ABB RobotStudio station: robot-studio-project.rspag

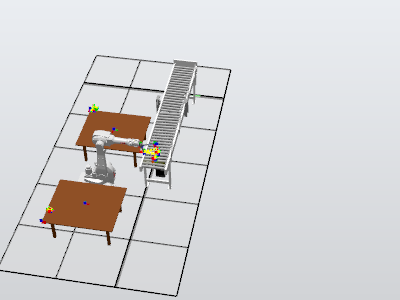
--- station ---
Station FinalConveyor (saved by RobotStudio 24.1.10693.0)
Controller IRB1600_6_145, task T_ROB1: task frame (RAPID world) sits at (2850, -850, 0) mm, rotated rx 0 ry 0 rz 90 deg in the station
Controller IRB1600_6_145
  mechanical unit ROB_1: IRB1600_6_145__03, 6 joints, base frame (0, 0, 0) mm
Layout (positions relative to the parent item):
  - big cube [part], size 200 x 200 x 200 mm
  - small cube [part], size 100 x 100 x 100 mm
  - Conveyor [smart component]
      signals: DI start_or_resume, DO cube_ready, DO cube_type
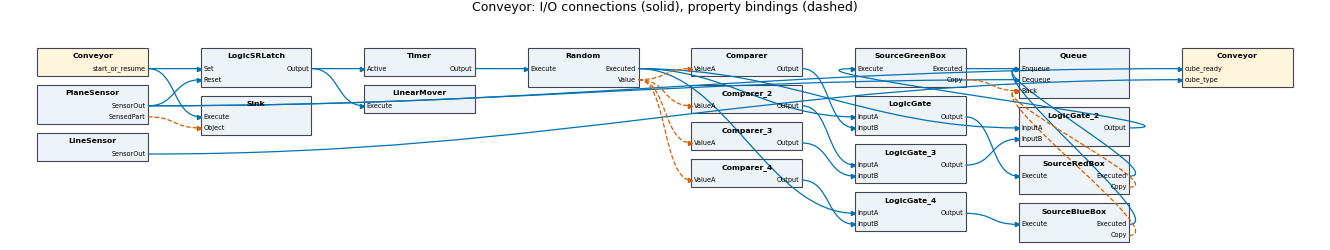
      connections:
        Timer.Output -> Random.Execute
        Random.Executed -> LogicGate.InputA
        Comparer.Output -> LogicGate.InputB
        Random.Executed -> LogicGate_2.InputA
        Comparer_2.Output -> LogicGate_3.InputA
        Comparer_3.Output -> LogicGate_3.InputB
        LogicGate_3.Output -> LogicGate_2.InputB
        Random.Executed -> LogicGate_4.InputA
        Comparer_4.Output -> LogicGate_4.InputB
        LogicGate.Output -> SourceRedBox.Execute
        LogicGate_2.Output -> SourceGreenBox.Execute
        LogicGate_4.Output -> SourceBlueBox.Execute
        SourceRedBox.Executed -> Queue.Enqueue
        SourceGreenBox.Executed -> Queue.Enqueue
        SourceBlueBox.Executed -> Queue.Enqueue
        Conveyor.start_or_resume -> LogicSRLatch.Set
        PlaneSensor.SensorOut -> Queue.Dequeue
        PlaneSensor.SensorOut -> LogicSRLatch.Reset
        LogicSRLatch.Output -> Timer.Active
        LogicSRLatch.Output -> LinearMover.Execute
        Conveyor.start_or_resume -> Sink.Execute
        PlaneSensor.SensorOut -> Conveyor.cube_ready
        LineSensor.SensorOut -> Conveyor.cube_type
        Random.Value => Comparer.ValueA
        Random.Value => Comparer_2.ValueA
        Random.Value => Comparer_3.ValueA
        Random.Value => Comparer_4.ValueA
        SourceRedBox.Copy => Queue.Back
        SourceGreenBox.Copy => Queue.Back
        SourceBlueBox.Copy => Queue.Back
        PlaneSensor.SensedPart => Sink.Object
    - SourceRedBox [smart component, from Components\Source.rslib]
        properties: Source=small cube; Copy=(none); Parent=(none); Position=[0.075 0.17 0.775]; Orientation=[0 0 0]; Transient=false; PhysicsBehavior=-1
    - SourceGreenBox [smart component, from Components\Source.rslib]
        properties: Source=small cube; Copy=(none); Parent=(none); Position=[0.075 0.17 0.775]; Orientation=[0 0 0]; Transient=false; PhysicsBehavior=-1
    - SourceBlueBox [smart component, from Components\Source.rslib]
        properties: Source=big cube; Copy=(none); Parent=(none); Position=[0.075 0.17 0.775]; Orientation=[0 0 0]; Transient=false; PhysicsBehavior=-1
    - Random [smart component, from Components\Random.rslib]
        properties: Value=1.86635471315419; Min=0; Max=3
    - Comparer [smart component, from Components\Comparer.rslib]
        properties: ValueA=1.86635471315419; Operator=<=; ValueB=1
    - Timer [smart component, from Components\Timer.rslib]
        properties: StartTime=0; Interval=2; Repeat=true; CurrentTime=0
    - Comparer_2 [smart component, from Components\Comparer.rslib]
        properties: ValueA=1.86635471315419; Operator=>; ValueB=1
    - Comparer_3 [smart component, from Components\Comparer.rslib]
        properties: ValueA=1.86635471315419; Operator=<=; ValueB=2
    - LogicGate [smart component, from Components\LogicGate.rslib]
        properties: Operator=AND; Delay=0
    - LogicGate_2 [smart component, from Components\LogicGate.rslib]
        properties: Operator=AND; Delay=0
    - LogicGate_3 [smart component, from Components\LogicGate.rslib]
        properties: Operator=AND; Delay=0
    - LogicGate_4 [smart component, from Components\LogicGate.rslib]
        properties: Operator=AND; Delay=0
    - Comparer_4 [smart component, from Components\Comparer.rslib]
        properties: ValueA=1.86635471315419; Operator=>; ValueB=2
    - Queue [smart component, from Components\Queue.rslib]
        properties: Back=(none); Front=(none); Queue={d5145b48-5921-41e5-a5cf-f289e25e2c56};{eb20e8fc-2243-4132-bafd-30e74f28caf8};{df543072-238f-4cf0-af28-d52d1ae9a375};{1c01fbfb-bd7a-479c-aabf-7e294c76dd45};{cb4fb4ea-8899-44f1-8836-deb4a8ef6429};{4a7ed11f-3483-4d0f-abfe-d523fadb1b42};{0f8e3dc3-db70-4297-9f91-4c7c364b3beb};{c87a5a8a-da50-415a-a569-0345de37618b};{a8b1a2bd-e0b2-4c05-9cb6-234d8fd6809a};{c18f4dcd-aaf8-47e2-ac1c-454d25c30403};{f1c64246-078b-4c03-92cf-52699b84a579};{05fd84a4-48ba-4786-b4e0-bb9a32800100};{2eff5ee7-084f-417a-bb43-7220eca7bcf1};{c83a14ee-1aed-4cfc-b806-602a5e6c2242};{0d87de5f-898c-47f1-911a-acb0e95ac153};{63b4051d-49dc-48c0-b256-ae6bb22b842a};{9f378025-0063-4114-8942-477e9b35e507};{4c7bcc95-1748-4e42-9dd8-063b71ec8c50};{8af862e1-0078-4417-b58c-83dbf2853366};{8bcf51d1-760d-4176-ac0d-77fba529ff68};{f84a91e3-2197-44a6-bd0c-9c5110243a1c};{99947171-f6ad-4ba1-92d8-702f21d52f91};{bc166aec-908d-47c2-b7d2-ad1fce975e4e}; NumberOfObjects=6
    - LinearMover [smart component, from Components\LinearMover.rslib]
        properties: Object=Queue; Direction=[1 0 0]; Speed=0.2; Reference=Global; ReferenceObject=(none)
    - PlaneSensor [smart component, from Components\PlaneSensor.rslib]
        properties: Origin=[2.910135 0.39 0.78]; Axis1=[0 -0.38 0]; Axis2=[0 0 0.1]; Tag=(none); SensedPart=(none)
      - _sensorPart_ [part], size 0 x 380 x 100 mm
    - LogicSRLatch [smart component, from Components\LogicSRLatch.rslib]
    - Sink [smart component, from Components\Sink.rslib]
        properties: Object=(none)
    - 400_guide [part], size 3033 x 590 x 945 mm
    - LineSensor [smart component, from Components\LineSensor.rslib]
        properties: Start=[2.8 0 0.95]; End=[2.8 0.3 0.95]; Length=0.3; Radius=0.001; Tag=(none); SensedPart=(none); SensedPoint=[0 0 0]
      - _sensorPart_ [part], size 2 x 300 x 2 mm
  - table_1 [part] at (2400, -1400, 500) mm, rotated rx 90 ry 0 rz 90 deg, size 1200 x 500 x 1000 mm
  - IRB1600_6_145__03 [mechanism] at (2850, -850, 0) mm, rotated rx 0 ry 0 rz 90 deg; joint values [0, 0, 0, 0, 0.5236, 0] (rad or m)
      links: Base, Link1, Link2, Link3, Link4, Link5, Link6
  - table_2 [part] at (4300, -1400, 500) mm, rotated rx 90 ry 0 rz 90 deg, size 1200 x 500 x 1000 mm
  - small cube test conveyor [part], size 100 x 100 x 100 mm
  - big cube test conveyor [part], size 200 x 200 x 200 mm
  - big cube test table [part], size 200 x 200 x 200 mm
  - small cube test table [part], size 100 x 100 x 100 mm
  - VacuumPenToolSC [smart component] at (2850, -43.71, 1154) mm, rotated rx 180 ry 60 rz -90 deg
      signals: DI diAttacher, DO doAttacher
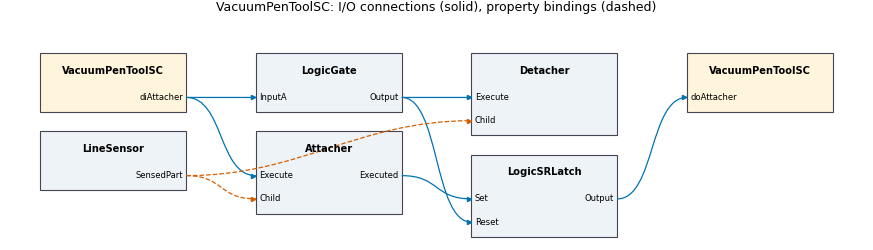
      connections:
        VacuumPenToolSC.diAttacher -> LogicGate.InputA
        LogicGate.Output -> Detacher.Execute
        Attacher.Executed -> LogicSRLatch.Set
        LogicSRLatch.Output -> VacuumPenToolSC.doAttacher
        VacuumPenToolSC.diAttacher -> Attacher.Execute
        LogicGate.Output -> LogicSRLatch.Reset
        LineSensor.SensedPart => Attacher.Child
        LineSensor.SensedPart => Detacher.Child
    - VacuumPenTool [mechanism] at (0, 0, 0) mm
        TCP VacuumTool at (106.34, 126.01, 0.37) mm, rotated rx -90 ry 0 rz -45 deg
        TCP PenTool at (-174.29, 194.28, 0.18) mm, rotated rx -90 ry 0 rz 45 deg
        links: DoubleToolVacuumPencil
    - LineSensor [smart component, from Components\LineSensor.rslib]
        properties: Start=[0.107 -0.00037 0.127]; End=[0.114 0 0.134]; Radius=0.001; SensedPart=(none); SensedPoint=[2.81016870117188 0.270228363037109 0.975]; Length=0.00990640701768306; Tag=(none)
      - _sensorPart_ [part], size 8.4 x 2.4 x 8.4 mm
    - Attacher [smart component, from Components\Attacher.rslib]
        properties: Parent=VacuumPenTool; Flange=0; Child=(none); Mount=false; Offset=[0 0 0]; Orientation=[0 0 0]
    - Detacher [smart component, from Components\Detacher.rslib]
        properties: Child=(none); KeepPosition=true
    - LogicGate [smart component, from Components\LogicGate.rslib]
        properties: Operator=NOT; Delay=0
    - LogicSRLatch [smart component, from Components\LogicSRLatch.rslib]
Attachment: VacuumPenToolSC is attached to IRB1600_6_145__03 / Link6
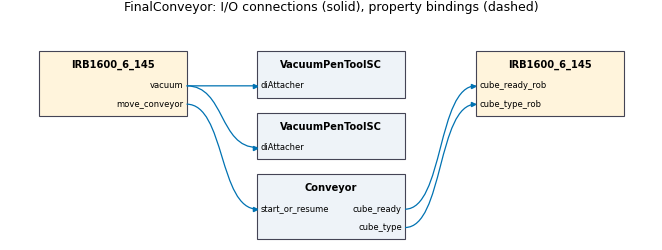
Station logic (signal -> signal, property => property):
  IRB1600_6_145.vacuum -> VacuumPenToolSC.diAttacher
  Conveyor.cube_ready -> IRB1600_6_145.cube_ready_rob
  Conveyor.cube_type -> IRB1600_6_145.cube_type_rob
  IRB1600_6_145.move_conveyor -> Conveyor.start_or_resume
  IRB1600_6_145.vacuum -> VacuumPenToolSC.diAttacher
Targets, tools, work objects and paths stored in the station and not in the controller backup, written as RAPID:
! task T_ROB1
MODULE Module1
  CONST robtarget pLocal:=[[0,0,0],[1,0,0,0],[0,0,0,0],[9E+09,9E+09,9E+09,9E+09,9E+09,9E+09]];
  PROC draw_big_cube()
    MoveJ Offs (bigcube_mid,0,0,-100),v200,z10,PenTool\WObj:=big_draw;
    MoveL Offs (bigcube_mid,50,50,0),v200,fine,PenTool\WObj:=big_draw;
    MoveL Offs (bigcube_mid,-50,-50,0),v50,fine,PenTool\WObj:=big_draw;
    MoveJ Offs (bigcube_mid,0,0,-100),v200,z10,PenTool\WObj:=big_draw;
  ENDPROC
  PROC draw_small_cube()
    MoveJ Offs (smallcube_mid,0,0,-50),v200,z10,PenTool\WObj:=small_draw;
    MoveL Offs (smallcube_mid,0,40,0),v200,fine,PenTool\WObj:=small_draw;
    MoveL Offs (smallcube_mid,0,-40,0),v50,fine,PenTool\WObj:=small_draw;
    MoveJ Offs (smallcube_mid,0,0,-50),v200,z10,PenTool\WObj:=small_draw;
  ENDPROC
ENDMODULE


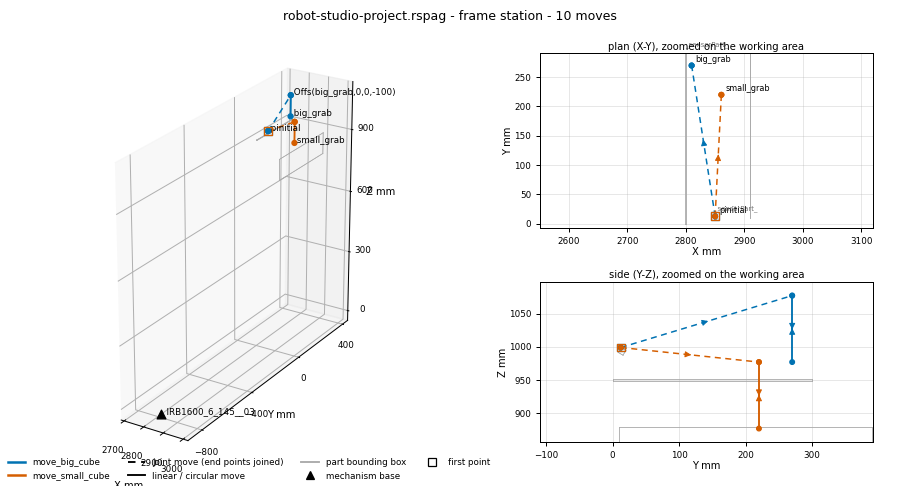
[picture p0: tool path of robot-studio-project.rspag in frame station, 10 of 25 moves have a stored position in this frame; points joined in program order, loops and branches not executed]
--- Controller Data/IRB1600_6_145/RAPID/TASK1/PROGMOD/CalibData.mod ---
MODULE CalibData
    PERS tooldata VacuumTool:=[TRUE,[[106.338,-0.37,126.015],[0.92388,0,0.382683,0]],[1,[0,0,1],[1,0,0,0],0,0,0]];
    PERS tooldata PenTool:=[TRUE,[[-174.289,-0.18,194.277],[0.92388,0,-0.382683,0]],[1,[0,0,1],[1,0,0,0],0,0,0]];
    TASK PERS wobjdata big_conveyor:=[FALSE,TRUE,"",[[1020,139.8,775],[0.707107,0,0,-0.707107]],[[100,100,200],[0,-0.707107,0.707107,0]]];
    TASK PERS wobjdata small_conveyor:=[FALSE,TRUE,"",[[1020,39,775],[0.707107,0,0,-0.707107]],[[50,50,100],[0,-0.707107,0.707107,0]]];
    TASK PERS wobjdata big_table:=[FALSE,TRUE,"",[[-550,1450,520],[0.707107,0,0,-0.707107]],[[500,600,0],[1,0,0,0]]];
    TASK PERS wobjdata big_draw:=[FALSE,TRUE,"",[[-550,1450,520],[0.707107,0,0,-0.707107]],[[200,150,200],[0,0,1,0]]];
    TASK PERS wobjdata small_table:=[FALSE,TRUE,"",[[-550,-1450,520],[1,0,0,0]],[[600,500,0],[1,0,0,0]]];
    TASK PERS wobjdata small_draw:=[FALSE,TRUE,"",[[-550,-1450,520],[1,0,0,0]],[[100,200,100],[0,-0.707107,0.707107,0]]];
ENDMODULE

--- Controller Data/IRB1600_6_145/RAPID/TASK1/PROGMOD/Module1.mod ---
MODULE Module1
    CONST robtarget pinitial:=[[862.254842504,-0.37,998.901090612],[0.130526193,0,0.991444861,0],[-1,0,-1,0],[9E+09,9E+09,9E+09,9E+09,9E+09,9E+09]];
    CONST robtarget big_grab:=[[0,0,-2],[1,0,0,0],[0,0,0,0],[9E+09,9E+09,9E+09,9E+09,9E+09,9E+09]];
    CONST robtarget big_release:=[[-300,-450,202],[0,1,0,0],[0,0,0,0],[9E+09,9E+09,9E+09,9E+09,9E+09,9E+09]];
    CONST robtarget small_grab:=[[0,0,-2],[1,0,0,0],[0,0,0,0],[9E+09,9E+09,9E+09,9E+09,9E+09,9E+09]];
    CONST robtarget small_release:=[[-500,-300,102],[0,0.707106781,0.707106781,0],[-2,0,-1,0],[9E+09,9E+09,9E+09,9E+09,9E+09,9E+09]];
    CONST robtarget bigcube_mid:=[[0,0,0],[1,0,0,0],[1,-1,-2,0],[9E+09,9E+09,9E+09,9E+09,9E+09,9E+09]];
    CONST robtarget smallcube_mid:=[[0,0,0],[1,0,0,0],[-2,0,1,0],[9E+09,9E+09,9E+09,9E+09,9E+09,9E+09]];

    VAR num layer_big := 0;
    VAR num row_big := 0;
    VAR num col_big := 0;

    VAR num layer_small := 0;
    VAR num row_small := 0;
    VAR num col_small := 0;

    PROC main()
        WHILE TRUE DO
            SetDO move_conveyor,1;
            WaitDI cube_ready_rob,1;
            SetDO move_conveyor,0;
            IF DInput(cube_type_rob) = 1 THEN
                IF row_big = 4 THEN
                    IF col_big = 2 THEN
                        row_big := 0;
                        col_big := 0;
                        layer_big := layer_big + 1;
                    ELSE
                        col_big := col_big + 1;
                        row_big := 0;
                    ENDIF
                ENDIF
                move_big_cube;
            ELSEIF DInput(cube_type_rob) = 0 THEN
                IF row_small = 6 THEN
                    IF col_small = 3 THEN
                        row_small := 0;
                        col_small := 0;
                        layer_small := layer_small + 1;
                    ELSE
                        col_small := col_small + 1;
                        row_small := 0;
                    ENDIF
                ENDIF
                move_small_cube;
            ENDIF
        ENDWHILE
    ENDPROC

    PROC move_big_cube()
        MoveJ pinitial,v1000,z100,VacuumTool\WObj:=wobj0;
        SetDO vacuum,0;
        MoveJ Offs(big_grab,0,0,-100),v500,z10,VacuumTool\WObj:=big_conveyor; !aproximation point above big cube in the conveyor
        MoveL big_grab,v50,fine,VacuumTool\WObj:=big_conveyor; !point to approach big cube
        WaitTime 1;
        SetDO vacuum,1;
        MoveL Offs(big_grab,0,0,-100),v200,z10,VacuumTool\WObj:=big_conveyor; !back to the aproximaton point
        MoveL Offs(big_release,300*col_big,300*row_big,50+200*layer_big),v1000,z100,VacuumTool\WObj:=big_table; !aproximation point above big cube in the table
        MoveL Offs(big_release,300*col_big,300*row_big,200*layer_big),v50,fine,VacuumTool\WObj:=big_table; !point to release big cube
        WaitTime 1;
        SetDO vacuum,0;
        MoveL Offs(big_release,300*col_big,300*row_big,50+200*layer_big),v1000,z100,VacuumTool\WObj:=big_table; !back to the aproximation point
        !draw 1,200;
        !MoveL Offs(big_release,300*col_big,300*row_big,50+200*layer_big),v1000,z100,VacuumTool\WObj:=big_table; !back to the aproximation point
        MoveL pinitial,v1000,z100,VacuumTool\WObj:=wobj0; !back to the initial point
        row_big := row_big + 1;
    ENDPROC

    PROC move_small_cube()
        MoveJ pinitial,v1000,z100,VacuumTool\WObj:=wobj0;
        SetDO vacuum,0;
        MoveJ Offs(small_grab,0,0,-100),v500,z10,VacuumTool\WObj:=small_conveyor; !aproximation point above small cube in the conveyor
        MoveL small_grab,v50,fine,VacuumTool\WObj:=small_conveyor; !point to approach small cube
        WaitTime 1;
        SetDO vacuum,1;
        MoveL Offs(small_grab,0,0,-100),v200,z10,VacuumTool\WObj:=small_conveyor; !back to the aproximaton point
        MoveL Offs(small_release,200*row_small,200*col_small,50+100*layer_small),v1000,z100,VacuumTool\WObj:=small_table; !aproximation point above small cube in the table
        MoveL Offs(small_release,200*row_small,200*col_small,100*layer_small),v50,fine,VacuumTool\WObj:=small_table; !point to release small cube
        WaitTime 1;
        SetDO vacuum,0;
        MoveL Offs(small_release,200*row_small,200*col_small,50+100*layer_small),v200,z100,VacuumTool\WObj:=small_table; !back to the aproximaton point
        draw 0,100;
        MoveL Offs(small_release,200*row_small,200*col_small,50+100*layer_small),v200,z100,VacuumTool\WObj:=small_table; !back to the aproximaton point
        MoveL pinitial,v1000,z100,VacuumTool\WObj:=wobj0; !back to the initial point
        row_small := row_small + 1;
    ENDPROC

    PROC draw(num type,num len)
        IF type = 1 THEN
            MoveJ Offs (bigcube_mid,300*col_big,-300*row_big,-len/2-200*layer_big),v200,z10,PenTool\WObj:=big_draw;
            MoveL Offs (bigcube_mid,300*col_big+len/4,len/4-300*row_big,-200*layer_big),v200,fine,PenTool\WObj:=big_draw;
            MoveL Offs (bigcube_mid,300*col_big-len/4,-len/4-300*row_big,-200*layer_big),v50,fine,PenTool\WObj:=big_draw;
            MoveJ Offs (bigcube_mid,300*col_big,-300*row_big,-len/2-200*layer_big),v200,z10,PenTool\WObj:=big_draw;
        ELSEIF type = 0 THEN
            MoveJ Offs (smallcube_mid,-200*col_small,-200*row_small,-len/2-100*layer_small),v200,z10,PenTool\WObj:=small_draw;
            MoveL Offs (smallcube_mid,-200*col_small,-len/4-200*row_small,-100*layer_small),v200,fine,PenTool\WObj:=small_draw;
            MoveL Offs (smallcube_mid,-200*col_small,len/4-200*row_small,-100*layer_small),v50,fine,PenTool\WObj:=small_draw;
            MoveJ Offs (smallcube_mid,-200*col_small,-200*row_small,-len/2-100*layer_small),v200,z10,PenTool\WObj:=small_draw;
        ENDIF
    ENDPROC

!    PROC draw_big_cube()
!        MoveJ Offs (bigcube_mid,0,0,-100),v200,z10,PenTool\WObj:=big_draw;
!        MoveL Offs (bigcube_mid,50,50,0),v200,fine,PenTool\WObj:=big_draw;
!        MoveL Offs (bigcube_mid,-50,-50,0),v50,fine,PenTool\WObj:=big_draw;
!        MoveJ Offs (bigcube_mid,0,0,-100),v200,z10,PenTool\WObj:=big_draw;
!    ENDPROC

!    PROC draw_small_cube()
!        MoveJ Offs (smallcube_mid,0,0,-50),v200,z10,PenTool\WObj:=small_draw;
!        MoveL Offs (smallcube_mid,0,40,0),v200,fine,PenTool\WObj:=small_draw;
!        MoveL Offs (smallcube_mid,0,-40,0),v50,fine,PenTool\WObj:=small_draw;
!        MoveJ Offs (smallcube_mid,0,0,-50),v200,z10,PenTool\WObj:=small_draw;
!    ENDPROC

ENDMODULE

--- Controller Data/IRB1600_6_145/SYSPAR/EIO.cfg ---
EIO:CFG_1.0:6:1::
#
EIO_SIGNAL:

      -Name "vacuum" -SignalType "DO"

      -Name "cube_ready_rob" -SignalType "DI"

      -Name "cube_type_rob" -SignalType "DI"

      -Name "move_conveyor" -SignalType "DO"
